PROGRAM VltFixtureCfc
VAR
END_VAR

END_PROGRAM

(* stored: Version 1.1.0.1, ProductVersion 3.1.4024.16
   POU VltFixtureCfc: Id {8aa4cfd7-a8c0-4d77-92fb-950ffec7d860}, SpecialFunc None *)
